// TIA Portal V20 export
// export: Created 2026-10-24T18:20:53.9485153Z, ExportSetting WithDefaults, DisplayName Totally Integrated Automation Portal, DisplayVersion V20 Update 6, DisplayName TIA Portal Openness, DisplayVersion V20 Update 6, DisplayName TIA Portal Version Control Interface, DisplayVersion V20 Update 6, DisplayName SINAMICS Startdrive Advanced, DisplayVersion V20 SP1 Update 2, DisplayName SINAMICS Startdrive G110M, G120, G120C, G120D, G120P, G115D, DisplayVersion V20 SP1 Update 2, DisplayName SINAMICS Startdrive G130, G150, S120, S150, SINAMICS MV, G220, S200, S210, DisplayVersion V20 SP1 Update 2, DisplayName STEP 7 Professional, DisplayVersion V20 Update 6, DisplayName STEP 7 Safety, DisplayVersion V20 Update 2, DisplayName WinCC Basic/Comfort/Advanced, DisplayVersion V20 Update 6, DisplayName WinCC Unified, DisplayVersion V20 Update 6
DATA_BLOCK "IDB_LadBoxes"   // DB2
VERSION : 0.1
// stored: AutoNumber true, DBAccessibleFromOPCUA true, DBAccessibleFromWebserver true, InstanceOfName FB_LadBoxes, InstanceOfType FB
"FB_LadBoxes"
   // VAR_INPUT
   //    Start : Bool;
   //    InValue : Int;
   //    Limit : Int;
   // END_VAR
   // VAR_OUTPUT
   //    Delayed : Bool;
   //    Copy : Int;
   //    Sum : Int;
   //    IsEqual : Bool;
   //    IsGreater : Bool;
   //    IsLessEqual : Bool;
   //    Average : Real;
   //    SectionsOk : Bool;
   //    Skipped : Bool;
   //    AfterJump : Bool;
   // END_VAR
   // VAR
   //    Delay { S7_SetPoint := 'True'} : TON_TIME;
   //    DelayElapsed : Time;
   //    Sections { S7_SetPoint := 'True'} : "FB_SclSections";
   //    Values : Array[0..9] of Real;
   //    SectionsBusy : Bool;
   //    SectionsSteps : Int;
   //    Setpoint : Real;
   // END_VAR
BEGIN
END_DATA_BLOCK
